(* IEC 61131-3 sources: SRCI_CLIENT_PLC/RobotLibrary/Library/POUs/Calculation/MC_LoadMeasurementAutomatic/Structures, 4 files *)

(* ---- LoadMeasurementAutomaticOutCmd.st ---- *)
{attribute 'pack_mode' := '1'}
// -------------------------------------------------------------------------
//  SRCI Robot Library
// -------------------------------------------------------------------------
//
//  Object:      LoadMeasurementAutomaticOutCmd
//  Author:      Thorsten Brach
//  Date:        2024-06-20
//
//  Description:
//
//
//  Copyright:
//    (C) 2024 Thorsten Brach. All rights reserved
//             Licensed under the MIT License.
//
//  Disclaimer:
//    This project is provided without any guarantee and can be used for
//    private and commercial purposes. Any use is at the user’s
//    own risk and responsibility.
//
// -------------------------------------------------------------------------
TYPE LoadMeasurementAutomaticOutCmd :
STRUCT
  /// FB is returning a unique ID for the cal led measurement.
  MeasuringID       : UINT;
  /// Measured load data (see chapter 5.5.6.4)
  LoadData          : LoadData;
  /// Load data available
  LoadDataAvailable : BOOL;
END_STRUCT
END_TYPE

(* ---- LoadMeasurementAutomaticParCmd.st ---- *)
{attribute 'pack_mode' := '1'}
// -------------------------------------------------------------------------
//  SRCI Robot Library
// -------------------------------------------------------------------------
//
//  Object:      LoadMeasurementAutomaticParCmd
//  Author:      Thorsten Brach
//  Date:        2024-06-20
//
//  Description:
//
//
//  Copyright:
//    (C) 2024 Thorsten Brach. All rights reserved
//             Licensed under the MIT License.
//
//  Disclaimer:
//    This project is provided without any guarantee and can be used for
//    private and commercial purposes. Any use is at the user’s
//    own risk and responsibility.
//
// -------------------------------------------------------------------------
TYPE LoadMeasurementAutomaticParCmd :
STRUCT
  /// Define which method should be used to measure the load data
  Mode               : LoadMeasurementMode;
  /// Define which mass is expected as a result of the load measurement
  Mass               : REAL;
  /// Define the area for the allowed motion of the Joint 3.
  /// The order of the two limit values does not matter.
  /// Only considered with "Mode" = 0, 2.
  Area_J3            : ARRAY[0..1] OF REAL;
  /// Define the area for the allowed motion of the Joint 4.
  /// The order of the two limit values does not matter.
  /// Only considered with "Mode" = 0, 2.
  Area_J4            : ARRAY[0..1] OF REAL;
  /// Define the area for the allowed motion of the Joint 5.
  /// The order of the two limit values does not matter.
  /// Only considered with "Mode" = 0, 2.
  Area_J5            : ARRAY[0..1] OF REAL;
  /// Define the area for the allowed motion of the Joint 6.
  /// The order of the two limit values does not matter.
  /// Only considered with "Mode" = 0, 2.
  Area_J6            : ARRAY[0..1] OF REAL;
  /// Define the first position for the load measurement.
  /// Only considered with "Mode" = 0, 1, 3 (ST-FIX F176: TWO_POSITIONS uses Position_1 and Position_2; the spec names 0, 1).
  Position_1         : RobotJointPosition;
  /// Define the second position for the load measurement.
  /// Only considered with "Mode" = 3.
  Position_2         : RobotJointPosition;
  /// Define the configuration angle for the load measurement.
  /// Only considered with "Mode" = 1.
  ConfigurationAngle : REAL;
END_STRUCT
END_TYPE

(* ---- LoadMeasurementAutomaticRecvData.st ---- *)
{attribute 'pack_mode' := '1'}
// -------------------------------------------------------------------------
//  SRCI Robot Library
// -------------------------------------------------------------------------
//
//  Object:      LoadMeasurementAutomaticRecvData
//  Author:      Thorsten Brach
//  Date:        2024-06-20
//
//  Description:
//
//
//  Copyright:
//    (C) 2024 Thorsten Brach. All rights reserved
//             Licensed under the MIT License.
//
//  Disclaimer:
//    This project is provided without any guarantee and can be used for
//    private and commercial purposes. Any use is at the user’s
//    own risk and responsibility.
//
// -------------------------------------------------------------------------
TYPE LoadMeasurementAutomaticRecvData EXTENDS RspHeader :
STRUCT
    /// FB is returning a unique ID for the cal led measurement.
  MeasuringID       : UINT;
  /// Measured load data (see chapter 5.5.6.4)
  LoadData          : LoadData;
  /// Load data available
  LoadDataAvailable : BOOL;
END_STRUCT
END_TYPE

(* ---- LoadMeasurementAutomaticSendData.st ---- *)
{attribute 'pack_mode' := '1'}
// -------------------------------------------------------------------------
//  SRCI Robot Library
// -------------------------------------------------------------------------
//
//  Object:      LoadMeasurementAutomaticSendData
//  Author:      Thorsten Brach
//  Date:        2024-06-20
//
//  Description:
//
//
//  Copyright:
//    (C) 2024 Thorsten Brach. All rights reserved
//             Licensed under the MIT License.
//
//  Disclaimer:
//    This project is provided without any guarantee and can be used for
//    private and commercial purposes. Any use is at the user’s
//    own risk and responsibility.
//
// -------------------------------------------------------------------------
TYPE LoadMeasurementAutomaticSendData EXTENDS CmdHeader:
STRUCT
    /// Define which mass is expected as a result of the load measurement
  Mass               : REAL;
  /// Define which method should be used to measure the load data
  Mode               : LoadMeasurementMode;
  /// Reserved
  Reserved           : BYTE;
  /// Define the area for the allowed motion of the Joint 3.
  /// The order of the two limit values does not matter.
  /// Only considered with "Mode" = 0, 2.
  Area_J3            : ARRAY[0..1] OF REAL;
  /// Define the area for the allowed motion of the Joint 4.
  /// The order of the two limit values does not matter.
  /// Only considered with "Mode" = 0, 2.
  Area_J4            : ARRAY[0..1] OF REAL;
  /// Define the area for the allowed motion of the Joint 5.
  /// The order of the two limit values does not matter.
  /// Only considered with "Mode" = 0, 2.
  Area_J5            : ARRAY[0..1] OF REAL;
  /// Define the area for the allowed motion of the Joint 6.
  /// The order of the two limit values does not matter.
  /// Only considered with "Mode" = 0, 2.
  Area_J6            : ARRAY[0..1] OF REAL;
  /// Define the configuration angle for the load measurement.
  /// Only considered with "Mode" = 1.
  ConfigurationAngle : REAL;
  /// Define the first position for the load measurement.
  /// Only considered with "Mode" = 0, 1.
  Position_1         : RobotJointPosition;
  /// Define the second position for the load measurement.
  /// Only considered with "Mode" = 3.
  Position_2         : RobotJointPosition;
END_STRUCT
END_TYPE
